// TIA Portal V20 export
// export: Created 2026-10-11T05:19:07.9521126Z, ExportSetting WithDefaults, DisplayName Totally Integrated Automation Portal, DisplayVersion V20, DisplayName TIA Portal Openness, DisplayVersion V20, DisplayName TIA Portal Teamcenter Gateway, DisplayVersion V20, DisplayName TIA Portal Version Control Interface, DisplayVersion V20, DisplayName SINAMICS Startdrive Advanced, DisplayVersion V20 SP1 Update 2, DisplayName SINAMICS Startdrive G110M, G120, G120C, G120D, G120P, G115D, DisplayVersion V20 SP1 Update 2, DisplayName SINAMICS Startdrive G130, G150, S120, S150, SINAMICS MV, G220, S200, S210, DisplayVersion V20 SP1 Update 2, DisplayName STEP 7 Professional, DisplayVersion V20, DisplayName STEP 7 Safety, DisplayVersion V20, DisplayName WinCC Basic/Comfort/Advanced, DisplayVersion V20, DisplayName WinCC Professional, DisplayVersion V20, DisplayName WinCC Unified, DisplayVersion V20
FUNCTION "FRK_ConfigUnit" : Void   // FC25, SCL
{ S7_Optimized_Access := 'TRUE' }
VERSION : 0.1
// stored: AutoNumber true, IsIECCheckEnabled false, SetENOAutomatically false, UDAEnableTagReadback false
   VAR_INPUT
      Scope : String;
      Policy : Array[0..6] of "ST_ModePolicy";
      ReadLevel : DInt;
      Readable : Bool;
   END_VAR
   VAR_IN_OUT
      Cursor : "FRK_ConfigCursor";
      Page : "ST_ConfigPage";
   END_VAR
   VAR_TEMP
      Index : Int;
      IndexText : String[8];
      Prefix : String[254];
      Item : String[254];
   END_VAR
BEGIN

   "FRK_ConfigAppend"(Scope := #Scope,
                      Item := 'CatalogCount',
                      ValueText := WSTRING#'0',
                      ValueType := 0,
                      ReadLevel := #ReadLevel,
                      Readable := #Readable,
                      Cursor := #Cursor,
                      Page := #Page);
   "FRK_ConfigAppend"(Scope := #Scope,
                      Item := 'AvailableModelCount',
                      ValueText := WSTRING#'0',
                      ValueType := 0,
                      ReadLevel := #ReadLevel,
                      Readable := #Readable,
                      Cursor := #Cursor,
                      Page := #Page);
   FOR #Index := 0 TO 6 DO
       #IndexText := INT_TO_STRING(#Index);
       IF #IndexText[1] = '+' THEN
           #IndexText := DELETE(IN := #IndexText, L := 1, P := 1);
       END_IF;
       #Prefix := CONCAT(IN1 := 'ModePolicy/ModePolicy[', IN2 := #IndexText);
       #Prefix := CONCAT(IN1 := #Prefix, IN2 := ']/');
       #Item := CONCAT(IN1 := #Prefix, IN2 := 'Shield');
       "FRK_ConfigAppend"(Scope := #Scope,
                          Item := #Item,
                          ValueText := STRING_TO_WSTRING(DINT_TO_STRING(#Policy[#Index].Shield)),
                          ValueType := 0,
                          ReadLevel := #ReadLevel,
                          Readable := #Readable,
                          Cursor := #Cursor,
                          Page := #Page);
       #Item := CONCAT(IN1 := #Prefix, IN2 := 'Style');
       "FRK_ConfigAppend"(Scope := #Scope,
                          Item := #Item,
                          ValueText := STRING_TO_WSTRING(DINT_TO_STRING(#Policy[#Index].Style)),
                          ValueType := 0,
                          ReadLevel := #ReadLevel,
                          Readable := #Readable,
                          Cursor := #Cursor,
                          Page := #Page);
   END_FOR;
END_FUNCTION
